{attribute 'Tc2GvlVarNames'}
VAR_GLOBAL
	(* Axis interface *)
	igGr05AxisClamp1			:AXIS_REF;							(* Interface plc -> nc *)

	(* Drive interface *)
	igGr05DriveClamp1			:ST_STOEBERSI6SC6CIA402_REF;		(* Interface nc -> plc *)

END_VAR

(* stored: Version 1.1.0.1, ProductVersion 3.1.4024.15
   GVL GVL_Gr05Interface: Id {89430459-3e23-4e74-97a8-bfdffe2a771e} *)
